FUNCTION_BLOCK FB_SboControlEnhanced EXTENDS FB_SboControl
VAR
END_VAR

METHOD Execute : BOOL
VAR
	bTestOk: BOOL; (*Used to cache the return value of the last '_OperativeTest' or '_DynamicTest' method call*)
	eError: E_AcsiServiceError; (*Used to cache the returned error of the last '_OperativeTest' or '_DynamicTest' method call*)
	tValue: T_UtcTime; (*Used to cache the current system time for 'tOpOk'*)
END_VAR
IF (_ipCtrl <> 0) AND_THEN (_ipCtrl.ipOper <> 0) THEN
	(* Initialize function block in the first cycle *)
	IF NOT bInit THEN
		_Init();
		bInit:=TRUE;
	END_IF

	CASE _eControlState OF
		E_SboControlState.Unselected:
			(* Check if ControlState changed in the last cycle *)
			IF bNewState THEN
				bNewState:=FALSE;
				_Reset();
			END_IF
			(* Check if a valid Cancel_req was received *)
			IF bCancelReq THEN
				bCancelReq:=FALSE;
			END_IF
			(* Check if a valid SelVal_req was received *)
			IF bSelValReq THEN
				bSelValReq:=FALSE;
				(* Go to next ControlState *)
				_eControlState:=E_SboControlState.Select_PerformTest;
				bNewState:=TRUE;
			END_IF

		E_SboControlState.Select_PerformTest:
			(* Check if ControlState changed in the last cycle *)
			IF bNewState THEN
				bNewState:=FALSE;
			END_IF
			(* Trigger the test until it is finished *)
			IF _Test(bTestOk=>bTestOk, eError=>eError) THEN
				IF bTestOk THEN
					(* Go to next ControlState *)
					_eControlState:=E_SboControlState.WaitForSelection;
				ELSE
					fbSelValCompletion.SetCompleted();
					fbSelValCompletion.eServiceError:=eError;
					(* Go back to ControlState 'Unselected' *)
					_eControlState:=E_SboControlState.Unselected;
				END_IF
				bNewState:=TRUE;
			END_IF

		E_SboControlState.WaitForSelection:
			(* Check if ControlState changed in the last cycle *)
			IF bNewState THEN
				bNewState:=FALSE;
			END_IF
			(* Set 'stSeld' *)
			IF (_ipCtrl.ipStSeld <> 0) THEN
				_ipCtrl.ipStSeld.bValue:=TRUE;
			END_IF
			fbSelValCompletion.SetCompleted();
			(* Go to next ControlState *)
			_eControlState:=E_SboControlState.Ready;
			bNewState:=TRUE;

		E_SboControlState.Ready:
			(* Check if ControlState changed in the last cycle *)
			IF bNewState THEN
				bNewState:=FALSE;
				(* Start timer *)
				IF (_ipCtrl.ipSboTimeout <> 0) THEN
					_fbSboTimer(IN:=TRUE, PT:=DWORD_TO_TIME(_ipCtrl.ipSboTimeout.nValue));
				END_IF
			END_IF
			_fbSboTimer();
			(* Check if a valid Cancel_req was received, 'sboTimeout' was exceeded or the association was lost *)
			IF bCancelReq OR_ELSE _fbSboTimer.Q OR_ELSE ((_ipCurrentAA <> 0) AND_THEN (_ipCurrentAA.eState <> E_AsyncEnvironmentState.Established)) THEN
				bCancelReq:=FALSE;
				_fbSboTimer(IN:=FALSE);
				(* Go to next ControlState *)
				_eControlState:=E_SboControlState.EndSelection;
				bNewState:=TRUE;
			END_IF
			(* Check if a valid Oper_req was received *)
			IF bOperReq THEN
				bOperReq:=FALSE;
				(* Go to next ControlState *)
				_eControlState:=E_SboControlState.PerformTest;
				bNewState:=TRUE;
			END_IF

		E_SboControlState.PerformTest:
			(* Check if ControlState changed in the last cycle *)
			IF bNewState THEN
				bNewState:=FALSE;
				(* Set 'opRcvd' *)
				IF (_ipCtrl.ipOpRcvd <> 0) THEN
					_ipCtrl.ipOpRcvd.bValue:=TRUE;
				END_IF
			END_IF
			(* Check if a valid Cancel_req was received *)
			IF bCancelReq THEN
				bCancelReq:=FALSE;
				(* Send Oper_resp- *)
				_SendLastApplError(ipAA:=_ipCurrentAA, ipCtrlData:=_ipCtrl.ipOper, eError:=E_AcsiApplError.NoError, ipOrigin:=_ipCtrl.ipOper.ipOrigin, ipCtlNum:=_ipCtrl.ipOper.ipCtlNum, eAddCause:=E_AcsiApplAddCause.AbortionByCancel);
				fbOperCompletion.SetCompleted();
				fbOperCompletion.eServiceError:=E_AcsiServiceError.AccessViolation;
				(* Go to ControlState 'EndSelection' *)
				_eControlState:=E_SboControlState.EndSelection;
				bNewState:=TRUE;
			END_IF
			(* Trigger the operative test until it is finished *)
			IF _OperativeTest(bOperativeTestOk=>bTestOk, eError=>eError) THEN
				(* Reset 'opRcvd' *)
				IF (_ipCtrl.ipOpRcvd <> 0) THEN
					_ipCtrl.ipOpRcvd.bValue:=FALSE;
				END_IF
				IF bTestOk THEN
					(* Go to next ControlState *)
					_eControlState:=E_SboControlState.WaitForExecution;
				ELSE
					fbOperCompletion.SetCompleted();
					fbOperCompletion.eServiceError:=eError;
					(* Go to ControlState 'EndSelection' *)
					_eControlState:=E_SboControlState.EndSelection;
				END_IF
				bNewState:=TRUE;
			END_IF

		E_SboControlState.WaitForExecution:
			(* Check if ControlState changed in the last cycle *)
			IF bNewState THEN
				bNewState:=FALSE;
			END_IF
			(* Check if a Cancel_req was received *)
			IF bCancelReq THEN
				bCancelReq:=FALSE;
				(* Send Oper_resp- *)
				_SendLastApplError(ipAA:=_ipCurrentAA, ipCtrlData:=_ipCtrl.ipOper, eError:=E_AcsiApplError.NoError, ipOrigin:=_ipCtrl.ipOper.ipOrigin, ipCtlNum:=_ipCtrl.ipOper.ipCtlNum, eAddCause:=E_AcsiApplAddCause.AbortionByCancel);
				fbOperCompletion.SetCompleted();
				fbOperCompletion.eServiceError:=E_AcsiServiceError.AccessViolation;
				(* Go to ControlState 'EndSelection' *)
				_eControlState:=E_SboControlState.EndSelection;
				bNewState:=TRUE;
			END_IF
			(* Trigger the dynamic test until it is finished *)
			IF _DynamicTest(bDynamicTestOk=>bTestOk, eError=>eError) THEN
				fbOperCompletion.SetCompleted();
				IF bTestOk THEN
					(* Go to next ControlState *)
					IF (_ipBehVal <> 0) AND_THEN ((_ipBehVal.eValue = E_AcsiBeh.TestBlocked) OR_ELSE (_ipBehVal.eValue = E_AcsiBeh.OnBlocked)) THEN
						_eControlState:=E_SboControlState.MirrorBlockedCommand;
					ELSE
						_eControlState:=E_SboControlState.WaitForChange;
					END_IF
				ELSE
					fbOperCompletion.eServiceError:=eError;
					(* Go to ControlState 'EndSelection' *)
					_eControlState:=E_SboControlState.EndSelection;
				END_IF
				bNewState:=TRUE;
			END_IF

		E_SboControlState.WaitForChange:
			(* Check if ControlState changed in the last cycle *)
			IF bNewState THEN
				bNewState:=FALSE;
				(* Set 'opOk' *)
				IF (_ipCtrl.ipOpOk <> 0) THEN
					_ipCtrl.ipOpOk.bValue:=TRUE;
				END_IF
				(* Set 'tOpOk' *)
				IF (_ipCtrl.ipTOpOk <> 0) AND_THEN (_ipCurrentAA <> 0) AND_THEN (_ipCurrentAA.GetSystemTime(tT=>tValue)) THEN
					_ipCtrl.ipTOpOk.tValue:=tValue;
				END_IF
			END_IF
			(* Update value *)
			_SetValue(uCtlVal:=_ipCtrl.ipOper.uCtlVal, ipCtlVal_AV:=_ipCtrl.ipOper.ipCtlVal_AnalogueValue);
			(* Update Timestamp 't' *)
			_UpdateTimestampValue(ipAA:=_ipCurrentAA);

			(* Reset 'opOk' *)
			IF (_ipCtrl.ipOpOk <> 0) THEN
				_ipCtrl.ipOpOk.bValue:=FALSE;
			END_IF
			(* Send CmdTerm_req+ *)
			_SendCommandTerminationReqPos(ipAA:=_ipCurrentAA, ipCtrlData:=_ipCtrl.ipOper);
			(* Go to next ControlState *)
			IF (_ipCtrl.ipSboClass <> 0) AND_THEN (_ipCtrl.ipSboClass.eValue = E_AcsiSboClasses.OperateMany) THEN
				_eControlState:=E_SboControlState.Ready;
			ELSE
				_eControlState:=E_SboControlState.EndSelection;
			END_IF
			bNewState:=TRUE;

		E_SboControlState.MirrorBlockedCommand:
			(* Check if ControlState changed in the last cycle *)
			IF bNewState THEN
				bNewState:=FALSE;
				(* Set 'opOk' *)
				IF (_ipCtrl.ipOpOk <> 0) THEN
					_ipCtrl.ipOpOk.bValue:=TRUE;
				END_IF
				(* Set 'tOpOk' *)
				IF (_ipCtrl.ipTOpOk <> 0) AND_THEN (_ipCurrentAA <> 0) AND_THEN (_ipCurrentAA.GetSystemTime(tT=>tValue)) THEN
					_ipCtrl.ipTOpOk.tValue:=tValue;
				END_IF
			END_IF
			(* Reset 'opOk' *)
			IF (_ipCtrl.ipOpOk <> 0) THEN
				_ipCtrl.ipOpOk.bValue:=FALSE;
			END_IF
			(* Send CmdTerm_req- *)
			_SendCommandTerminationReqNeg(ipAA:=_ipCurrentAA, ipCtrlData:=_ipCtrl.ipOper, eError:=E_AcsiApplError.NoError, ipOrigin:=_ipCtrl.ipOper.ipOrigin, ipCtlNum:=_ipCtrl.ipOper.ipCtlNum, eAddCause:=E_AcsiApplAddCause.BlockedByMode);
			(* Go to next ControlState *)
			IF (_ipCtrl.ipSboClass <> 0) AND_THEN (_ipCtrl.ipSboClass.eValue = E_AcsiSboClasses.OperateMany) THEN
				_eControlState:=E_SboControlState.Ready;
			ELSE
				_eControlState:=E_SboControlState.EndSelection;
			END_IF
			bNewState:=TRUE;

		E_SboControlState.EndSelection:
			(* Check if ControlState changed in the last cycle *)
			IF bNewState THEN
				bNewState:=FALSE;
				(* Reset 'stSeld' *)
				IF (_ipCtrl.ipStSeld <> 0) THEN
					_ipCtrl.ipStSeld.bValue:=FALSE;
				END_IF
			END_IF
			(* Go to next ControlState *)
			_eControlState:=E_SboControlState.Unselected;
			bNewState:=TRUE;
	END_CASE
END_IF

(* Monitor transmission of LastApplError *)
CASE _nLastApplErrorReqState OF
	0:	;
	1:
		IF (_ipLastApplErrorReq <> 0) THEN
			Execute:=_ipLastApplErrorReq.Execute();
			IF NOT _ipLastApplErrorReq.IsBusy() THEN
				IF _ipLastApplErrorReq.IsCompleted() THEN
					SUPER^.SetCompleted();
				ELSE
					SUPER^.CopyFrom(ipSource:=_ipLastApplErrorReq);
				END_IF
				_nLastApplErrorReqState:=0;
			END_IF
		END_IF
END_CASE
(* Monitor transmission of CommandTermination *)
CASE _nCmdTermReqState OF
	0:	RETURN;
	1:
		IF (_ipCmdTermReq <> 0) THEN
			Execute:=_ipCmdTermReq.Execute();
			IF NOT _ipCmdTermReq.IsBusy() THEN
				IF _ipCmdTermReq.IsCompleted() THEN
					SUPER^.SetCompleted();
				ELSE
					SUPER^.CopyFrom(ipSource:=_ipLastApplErrorReq);
				END_IF
				_nCmdTermReqState:=0;
			END_IF
		END_IF
END_CASE
END_METHOD

METHOD OnCompletionWaitEvent : BOOL
VAR_INPUT
	ipDai: I_AcsiDataAccessInfoClass;
	ipData: I_AcsiCommonDataClass;
	eFc: E_AcsiFc;
END_VAR
VAR_OUTPUT
	ipResult: I_AcsiServiceResultClass := fbCompletion;
END_VAR
VAR
	eServiceError: E_AcsiServiceError;
	ipAA: I_ScsmAssociationClass; (*Interface pointer to application association*)
END_VAR
fbCompletion.SetCompleted();
IF (ipDai = 0) OR_ELSE (ipData = 0) THEN
	fbCompletion.eServiceError:=E_AcsiServiceError.AccessViolation;
	RETURN;
END_IF

(* Check if an Operate request is received *)
IF (ipDai.eService = E_AcsiServiceType.SetDataValues) THEN
	IF	(ipData.sObjectName = 'Oper') THEN
		fbOperCompletion.SetBusy();
		ipResult:=fbOperCompletion;
		bOperReq:=TRUE;
		OnCompletionWaitEvent:=TRUE;
	ELSIF (ipData.sObjectName = 'SBOw') THEN
		ScsmAssociation_From_Dai(in:=ipDai, out=>_ipCurrentAA);
		fbSelValCompletion.SetBusy();
		ipResult:=fbSelValCompletion;
		bSelValReq:=TRUE;
		OnCompletionWaitEvent:=TRUE;
	ELSIF (ipData.sObjectName = 'Cancel') THEN
		fbCancelCompletion.SetCompleted();
		ipResult:=fbCancelCompletion;
		IF _CheckCancelReq(ipDai:=ipDai, eError=>eServiceError) THEN
			bCancelReq:=TRUE;
		ELSE
			fbCancelCompletion.eServiceError:=eServiceError;
		END_IF
	END_IF
END_IF
END_METHOD

(*Implementation of user application data update event method.*)
METHOD OnGetVEvent
VAR_INPUT
	ipDai: I_AcsiDataAccessInfoClass; (*Additional data access info*)
	ipData: I_AcsiCommonDataClass; (*Interface pointer to data object*)
	eFc: E_AcsiFc; (*Functional constraint*)
END_VAR
VAR
END_VAR
END_METHOD

(*Implementation of user application data update event method.*)
METHOD OnGetVPreEvent : E_AcsiServiceError
VAR_INPUT
	ipDai: I_AcsiDataAccessInfoClass; (*Additional data access info*)
	ipData: I_AcsiCommonDataClass; (*Interface pointer to data object*)
	eFc: E_AcsiFc; (*Functional constraint*)
END_VAR
VAR
END_VAR
END_METHOD

(*Implementation of user application data update event method.*)
METHOD OnSetVPreEvent : E_AcsiServiceError
VAR_INPUT
	ipDai: I_AcsiDataAccessInfoClass; (*Additional data access info*)
	ipMemory: I_AnyMemoryBuffer; (*Interface pointer to buffer containig new value data*)
	ipData: I_AcsiCommonDataClass; (*Interface pointer to data object*)
	eFc: E_AcsiFc; (*Functional constraint*)
END_VAR
VAR_OUTPUT
	ipLastApplError: I_AcsiDATypeLastApplError; (*IF <> 0 => send LastApplError request*)
END_VAR
VAR
	ipAA: I_ScsmAssociationClass; (*Interface pointer to application association*)
	bItself: BOOL; (*If TRUE => Checking object is sub-data object itself*)
END_VAR
IF (eFc = E_AcsiFc.CO) AND_THEN (_ipCtrl <> 0) AND_THEN (ipDai <> 0) AND_THEN (ipDai.Write) AND_THEN (ipDai.ipAccessData <> 0) AND_THEN (ipData <> 0)
AND_THEN ScsmAssociation_From_Dai(in:=ipDai, out=>ipAA) THEN
	IF (_ipCtrl.ipOper <> 0) AND_THEN (_ipCtrl.ipOper.ipOrigin <> 0) AND_THEN (_ipCtrl.ipOper.ipCtlNum <> 0) THEN
		(* Check for invalid write attemps to prevent 'Oper' from being overwritten while a control request is being executed *)
		IF (ipDai.ipAccessData.sObjectName = 'Oper') THEN
			(* Only allow 'Oper' requests in state 'Ready' *)
			IF (_eControlState <> E_SboControlState.Ready) THEN
				ipLastApplError:=ipAA.SetAdditionalCauseDiag(ipCtrlData:=_ipCtrl.ipOper, eError:=E_AcsiApplError.NoError, stOrigin:=_ipCtrl.ipOper.ipOrigin.stOrigin, nCtlNum:=_ipCtrl.ipOper.ipCtlNum.nValue, eAddCause:=E_AcsiApplAddCause.CommandAlreadyInExecution);
				OnSetVPreEvent:=E_AcsiServiceError.AccessViolation;
				RETURN;
			END_IF
		ELSIF (_ipCtrl.ipOper.HasDataSubObject(ipData:=ipDai.ipAccessData, bItself=>bItself) AND_THEN (NOT bItself)) THEN
			(* Don't allow write access to subdata of 'Oper'*)
			ipLastApplError:=ipAA.SetAdditionalCauseDiag(ipCtrlData:=_ipCtrl.ipOper, eError:=E_AcsiApplError.NoError, stOrigin:=_ipCtrl.ipOper.ipOrigin.stOrigin, nCtlNum:=_ipCtrl.ipOper.ipCtlNum.nValue, eAddCause:=E_AcsiApplAddCause.NotSupported);
			OnSetVPreEvent:=E_AcsiServiceError.AccessViolation;
			RETURN;
		END_IF
	END_IF
	IF (_ipCtrl.ipSBOw <> 0) AND_THEN (_ipCtrl.ipSBOw.ipOrigin <> 0) AND_THEN (_ipCtrl.ipSBOw.ipCtlNum <> 0) THEN
		(* Check for invalid write attemps to prevent 'SBOw' from being overwritten while a control request is being executed *)
		IF (ipDai.ipAccessData.sObjectName = 'SBOw') THEN
			(* Only allow 'SelectWithValue' requests in state 'Unselected' *)
			IF (_eControlState <> E_SboControlState.Unselected) THEN
				ipLastApplError:=ipAA.SetAdditionalCauseDiag(ipCtrlData:=_ipCtrl.ipSBOw, eError:=E_AcsiApplError.NoError, stOrigin:=_ipCtrl.ipSBOw.ipOrigin.stOrigin, nCtlNum:=_ipCtrl.ipSBOw.ipCtlNum.nValue, eAddCause:=E_AcsiApplAddCause.CommandAlreadyInExecution);
				OnSetVPreEvent:=E_AcsiServiceError.AccessViolation;
				RETURN;
			ELSIF (_ipCtrl.ipSBOw.HasDataSubObject(ipData:=ipDai.ipAccessData, bItself=>bItself) AND_THEN (NOT bItself)) THEN
				(* Don't allow write access to subdata of 'SBOw'*)
				ipLastApplError:=ipAA.SetAdditionalCauseDiag(ipCtrlData:=_ipCtrl.ipSBOw, eError:=E_AcsiApplError.NoError, stOrigin:=_ipCtrl.ipSBOw.ipOrigin.stOrigin, nCtlNum:=_ipCtrl.ipSBOw.ipCtlNum.nValue, eAddCause:=E_AcsiApplAddCause.NotSupported);
				OnSetVPreEvent:=E_AcsiServiceError.AccessViolation;
				RETURN;
			END_IF
		END_IF
	END_IF
	IF (_ipCtrl.ipCancel <> 0) AND_THEN (_ipCtrl.ipCancel.ipOrigin <> 0) AND_THEN (_ipCtrl.ipCancel.ipCtlNum <> 0) THEN
		IF (ipDai.ipAccessData.sObjectName <> 'Cancel') AND_THEN (_ipCtrl.ipCancel.HasDataSubObject(ipData:=ipDai.ipAccessData)) THEN
			(* Don't allow write access to subdata of 'Cancel'*)
			ipLastApplError:=ipAA.SetAdditionalCauseDiag(ipCtrlData:=_ipCtrl.ipCancel, eError:=E_AcsiApplError.NoError, stOrigin:=_ipCtrl.ipCancel.ipOrigin.stOrigin, nCtlNum:=_ipCtrl.ipCancel.ipCtlNum.nValue, eAddCause:=E_AcsiApplAddCause.NotSupported);
			OnSetVPreEvent:=E_AcsiServiceError.AccessViolation;
			RETURN;
		END_IF
	END_IF
END_IF
END_METHOD

END_FUNCTION_BLOCK

(* stored: Version 1.1.0.1
   POU FB_SboControlEnhanced: Id {989b00d1-db0f-4d85-b079-231a7ae28e8c}, SpecialFunc None
   Method Execute: Id {7123b31b-40df-4c06-bdc6-5323d479de3d}
   Method OnCompletionWaitEvent: Id {8f733670-1e0f-4c54-a57c-3a62f75ecc2a}
   Method OnGetVEvent: Id {af81ec72-660c-44ce-ab42-22fdf5c75a15}
   Method OnGetVPreEvent: Id {cd5c264c-f01f-48a9-91f0-98bde6b4164d}
   Method OnSetVPreEvent: Id {00160a85-f639-488d-b191-3e1c80123df6} *)
